# EPICS substitutions: iocs/motor/aerotech-ioc/db/Soloist.substitutions
# C's iocAerotech Soloist.substitutions, P from st.cmd.
file "$(MOTOR)/db/motor.db"
{
pattern
{N,  M,       DTYP,       C,  S,  DESC,          EGU,      DIR,  VELO,  VBAS,  ACCL,  BDST,  BVEL,  BACC,  MRES,    PREC,  DHLM,  DLLM,  INIT}
{2,  "m$(N)", "Soloist",  0,  0,  "motor $(N)",  degrees,  Pos,  1,     .1,    .2,    0,     1,     .2,    2.5e-4,  5,     100,   -100,  ""}
}
